// TIA Portal V20 export
// export: Created 2026-10-19T18:07:30.6086494Z, ExportSetting WithDefaults, DisplayName Totally Integrated Automation Portal, DisplayVersion V20 Update 6, DisplayName TIA Portal Openness, DisplayVersion V20 Update 6, DisplayName TIA Portal Version Control Interface, DisplayVersion V20 Update 6, DisplayName SINAMICS Startdrive Advanced, DisplayVersion V20 SP1, DisplayName SINAMICS Startdrive G130, G150, S120, S150, SINAMICS MV, G220, S200, S210, DisplayVersion V20 SP1, DisplayName SINAMICS Startdrive G110M, G120, G120C, G120D, G120P, G115D, DisplayVersion V20 SP1, DisplayName STEP 7 Professional, DisplayVersion V20 Update 6, DisplayName STEP 7 Safety, DisplayVersion V20 Update 2, DisplayName WinCC Basic/Comfort/Advanced, DisplayVersion V20 Update 6, DisplayName WinCC Unified, DisplayVersion V20 Update 6
FUNCTION_BLOCK "SICK_Barcode_FB"   // FB19, SCL
{ S7_Optimized_Access := 'TRUE' }
VERSION : 0.1
// stored: AutoNumber true, IsIECCheckEnabled false, IsRetainMemResEnabled false, MemoryReserve 100, SetENOAutomatically false, UDAEnableTagReadback false
   VAR_INPUT
      Rd_Done : Bool;
      Req_Done : Bool;
      Req_Busy : Bool;
      Error : Bool;
      arrResult : Array[1..200] of Byte;
      iCounter : USInt;
      iLength : Int;
      Error_Code : DWord;
   END_VAR
   VAR_OUTPUT
      Test_Comm : Bool;
      Enable_Trigger : Bool;
      Disable_Trigger : Bool;
      Enable_Req : Bool;
      Result : String;
      Test_OK : Bool;
   END_VAR
BEGIN
   //Communication Test
   IF "VTD_BCD_Start_Comm_Test_HMI_Tag" THEN
       #Test_Comm := 1;
       #Enable_Req := 1;
       "IEC_Timer_0_DB_1".TON(IN:=True,
                              PT:=t#1s);
   END_IF;

   //TEST OK
   IF #Req_Done AND "IEC_Timer_0_DB_1".Q AND NOT #Error THEN
       #Test_OK := 1;
       #Test_Comm := 0;
       #Enable_Req := 0;
       "VTD_BCD_Start_Comm_Test_HMI_Tag" := 0;
       "IEC_Timer_0_DB_1".TON(IN := FALSE,
                              PT := t#0s);
   END_IF;

   //ERROR
   IF "IEC_Timer_0_DB_1".Q AND #Error THEN
           #Test_OK := 0;
           #Test_Comm := 0;
           #Enable_Req := 0;
           "VTD_BCD_Start_Comm_Test_HMI_Tag" := 0;
           "IEC_Timer_0_DB_1".TON(IN := FALSE,
                                  PT := t#0s);
       END_IF;

   //Enable Trigger
       IF "VTD_BCD_Enable_Trigger_HMI_Tag" OR "Auto_Start_Barcode" THEN
       #Enable_Trigger := 1;
       #Enable_Req := 1;
       "VTD_BCD_Disable_Trigger_HMI_Tag" := 0;
       #Disable_Trigger := 0;
   //Disable Trigger
   ELSIF "VTD_BCD_Disable_Trigger_HMI_Tag" OR "Auto_Stop_Barcode" THEN
       #Disable_Trigger := 1;
       #Enable_Req := 1;
       "VTD_BCD_Enable_Trigger_HMI_Tag" := 0;
       #Enable_Trigger := 0;
   ELSE
       #Enable_Trigger := 0;
       #Enable_Req := 0;
       #Disable_Trigger := 0;
   END_IF;


   "R_TRIG_DB_5"(CLK:=#Rd_Done);

   IF "R_TRIG_DB_5".Q OR "IEC_Timer_0_DB_18".Q OR
       ("VTD_BCD_Enable_Trigger_HMI_Tag" AND "VTD_BCD_Disable_Trigger_HMI_Tag")
   THEN
       "VTD_BCD_Disable_Trigger_HMI_Tag" := 0;
       #Enable_Trigger := 0;
       #Disable_Trigger := 0;
       #Enable_Req := 0;
       "IEC_Timer_0_DB_18".TON(IN := FALSE,
                               PT := T#0S);
       "Auto_Stop_Barcode" := 0;
   END_IF;

   "IEC_Timer_0_DB_18".TON(IN:=("VTD_BCD_Enable_Trigger_HMI_Tag" OR "VTD_BCD_Disable_Trigger_HMI_Tag" OR "Auto_Start_Barcode" OR "Auto_Stop_Barcode"),
                               PT:=T#10S);

   #Result := "ByteArrayToString_1"(Lenght := #iLength, ByteArray := #arrResult);
END_FUNCTION_BLOCK
